Staubli VAL3: onSimulate.pgx

public program onSimulate()
begin
end
